IF SUPER^.Step(981,TRUE,'Step number 981') THEN		
	SUPER^.StepCompleteWhen((_runOneStep OR _runAllSteps) AND _finishStep);	
	IF _runOneStep THEN	
		_runOneStep := FALSE;
		RETURN;
	END_IF	
END_IF		
		
IF SUPER^.Step(982,TRUE,'Step number 982') THEN		
	SUPER^.StepCompleteWhen((_runOneStep OR _runAllSteps) AND _finishStep);	
	IF _runOneStep THEN	
		_runOneStep := FALSE;
		RETURN;
	END_IF	
END_IF		
		
IF SUPER^.Step(983,TRUE,'Step number 983') THEN		
	SUPER^.StepCompleteWhen((_runOneStep OR _runAllSteps) AND _finishStep);	
	IF _runOneStep THEN	
		_runOneStep := FALSE;
		RETURN;
	END_IF	
END_IF		
		
IF SUPER^.Step(984,TRUE,'Step number 984') THEN		
	SUPER^.StepCompleteWhen((_runOneStep OR _runAllSteps) AND _finishStep);	
	IF _runOneStep THEN	
		_runOneStep := FALSE;
		RETURN;
	END_IF	
END_IF		
		
IF SUPER^.Step(985,TRUE,'Step number 985') THEN		
	SUPER^.StepCompleteWhen((_runOneStep OR _runAllSteps) AND _finishStep);	
	IF _runOneStep THEN	
		_runOneStep := FALSE;
		RETURN;
	END_IF	
END_IF		
		
IF SUPER^.Step(986,TRUE,'Step number 986') THEN		
	SUPER^.StepCompleteWhen((_runOneStep OR _runAllSteps) AND _finishStep);	
	IF _runOneStep THEN	
		_runOneStep := FALSE;
		RETURN;
	END_IF	
END_IF		
		
IF SUPER^.Step(987,TRUE,'Step number 987') THEN		
	SUPER^.StepCompleteWhen((_runOneStep OR _runAllSteps) AND _finishStep);	
	IF _runOneStep THEN	
		_runOneStep := FALSE;
		RETURN;
	END_IF	
END_IF		
		
IF SUPER^.Step(988,TRUE,'Step number 988') THEN		
	SUPER^.StepCompleteWhen((_runOneStep OR _runAllSteps) AND _finishStep);	
	IF _runOneStep THEN	
		_runOneStep := FALSE;
		RETURN;
	END_IF	
END_IF		
		
IF SUPER^.Step(989,TRUE,'Step number 989') THEN		
	SUPER^.StepCompleteWhen((_runOneStep OR _runAllSteps) AND _finishStep);	
	IF _runOneStep THEN	
		_runOneStep := FALSE;
		RETURN;
	END_IF	
END_IF		
		
IF SUPER^.Step(990,TRUE,'Step number 990') THEN		
	SUPER^.StepCompleteWhen((_runOneStep OR _runAllSteps) AND _finishStep);	
	IF _runOneStep THEN	
		_runOneStep := FALSE;
		RETURN;
	END_IF	
END_IF		
		
IF SUPER^.Step(991,TRUE,'Step number 991') THEN		
	SUPER^.StepCompleteWhen((_runOneStep OR _runAllSteps) AND _finishStep);	
	IF _runOneStep THEN	
		_runOneStep := FALSE;
		RETURN;
	END_IF	
END_IF		
		
IF SUPER^.Step(992,TRUE,'Step number 992') THEN		
	SUPER^.StepCompleteWhen((_runOneStep OR _runAllSteps) AND _finishStep);	
	IF _runOneStep THEN	
		_runOneStep := FALSE;
		RETURN;
	END_IF	
END_IF		
		
IF SUPER^.Step(993,TRUE,'Step number 993') THEN		
	SUPER^.StepCompleteWhen((_runOneStep OR _runAllSteps) AND _finishStep);	
	IF _runOneStep THEN	
		_runOneStep := FALSE;
		RETURN;
	END_IF	
END_IF		
		
IF SUPER^.Step(994,TRUE,'Step number 994') THEN		
	SUPER^.StepCompleteWhen((_runOneStep OR _runAllSteps) AND _finishStep);	
	IF _runOneStep THEN	
		_runOneStep := FALSE;
		RETURN;
	END_IF	
END_IF		
		
IF SUPER^.Step(995,TRUE,'Step number 995') THEN		
	SUPER^.StepCompleteWhen((_runOneStep OR _runAllSteps) AND _finishStep);	
	IF _runOneStep THEN	
		_runOneStep := FALSE;
		RETURN;
	END_IF	
END_IF		
		
IF SUPER^.Step(996,TRUE,'Step number 996') THEN		
	SUPER^.StepCompleteWhen((_runOneStep OR _runAllSteps) AND _finishStep);	
	IF _runOneStep THEN	
		_runOneStep := FALSE;
		RETURN;
	END_IF	
END_IF		
		
IF SUPER^.Step(997,TRUE,'Step number 997') THEN		
	SUPER^.StepCompleteWhen((_runOneStep OR _runAllSteps) AND _finishStep);	
	IF _runOneStep THEN	
		_runOneStep := FALSE;
		RETURN;
	END_IF	
END_IF		
		
IF SUPER^.Step(998,TRUE,'Step number 998') THEN		
	SUPER^.StepCompleteWhen((_runOneStep OR _runAllSteps) AND _finishStep);	
	IF _runOneStep THEN	
		_runOneStep := FALSE;
		RETURN;
	END_IF	
END_IF		
		
IF SUPER^.Step(999,TRUE,'Step number 999') THEN		
	SUPER^.StepCompleteWhen((_runOneStep OR _runAllSteps) AND _finishStep);	
	IF _runOneStep THEN	
		_runOneStep := FALSE;
		RETURN;
	END_IF	
END_IF		
		
IF SUPER^.Step(1000,TRUE,'Step number 1000') THEN		
	SUPER^.StepCompleteWhen((_runOneStep OR _runAllSteps) AND _finishStep);	
	IF _runOneStep THEN	
		_runOneStep := FALSE;
		RETURN;
	END_IF	
END_IF		
		
IF SUPER^.Step(1001,TRUE,'Step number 1001') THEN		
	SUPER^.StepCompleteWhen((_runOneStep OR _runAllSteps) AND _finishStep);	
	IF _runOneStep THEN	
		_runOneStep := FALSE;
		RETURN;
	END_IF	
END_IF		
		
IF SUPER^.Step(1002,TRUE,'Step number 1002') THEN		
	SUPER^.StepCompleteWhen((_runOneStep OR _runAllSteps) AND _finishStep);	
	IF _runOneStep THEN	
		_runOneStep := FALSE;
		RETURN;
	END_IF	
END_IF		
		
IF SUPER^.Step(1003,TRUE,'Step number 1003') THEN		
	SUPER^.StepCompleteWhen((_runOneStep OR _runAllSteps) AND _finishStep);	
	IF _runOneStep THEN	
		_runOneStep := FALSE;
		RETURN;
	END_IF	
END_IF		
		
IF SUPER^.Step(1004,TRUE,'Step number 1004') THEN		
	SUPER^.StepCompleteWhen((_runOneStep OR _runAllSteps) AND _finishStep);	
	IF _runOneStep THEN	
		_runOneStep := FALSE;
		RETURN;
	END_IF	
END_IF		
		
IF SUPER^.Step(1005,TRUE,'Step number 1005') THEN		
	SUPER^.StepCompleteWhen((_runOneStep OR _runAllSteps) AND _finishStep);	
	IF _runOneStep THEN	
		_runOneStep := FALSE;
		RETURN;
	END_IF	
END_IF		
		
IF SUPER^.Step(1006,TRUE,'Step number 1006') THEN		
	SUPER^.StepCompleteWhen((_runOneStep OR _runAllSteps) AND _finishStep);	
	IF _runOneStep THEN	
		_runOneStep := FALSE;
		RETURN;
	END_IF	
END_IF		
		
IF SUPER^.Step(1007,TRUE,'Step number 1007') THEN		
	SUPER^.StepCompleteWhen((_runOneStep OR _runAllSteps) AND _finishStep);	
	IF _runOneStep THEN	
		_runOneStep := FALSE;
		RETURN;
	END_IF	
END_IF		
		
IF SUPER^.Step(1008,TRUE,'Step number 1008') THEN		
	SUPER^.StepCompleteWhen((_runOneStep OR _runAllSteps) AND _finishStep);	
	IF _runOneStep THEN	
		_runOneStep := FALSE;
		RETURN;
	END_IF	
END_IF		
		
IF SUPER^.Step(1009,TRUE,'Step number 1009') THEN		
	SUPER^.StepCompleteWhen((_runOneStep OR _runAllSteps) AND _finishStep);	
	IF _runOneStep THEN	
		_runOneStep := FALSE;
		RETURN;
	END_IF	
END_IF		
		
IF SUPER^.Step(1010,TRUE,'Step number 1010') THEN		
	SUPER^.StepCompleteWhen((_runOneStep OR _runAllSteps) AND _finishStep);	
	IF _runOneStep THEN	
		_runOneStep := FALSE;
		RETURN;
	END_IF	
END_IF		
		
IF SUPER^.Step(1011,TRUE,'Step number 1011') THEN		
	SUPER^.StepCompleteWhen((_runOneStep OR _runAllSteps) AND _finishStep);	
	IF _runOneStep THEN	
		_runOneStep := FALSE;
		RETURN;
	END_IF	
END_IF		
		
IF SUPER^.Step(1012,TRUE,'Step number 1012') THEN		
	SUPER^.StepCompleteWhen((_runOneStep OR _runAllSteps) AND _finishStep);	
	IF _runOneStep THEN	
		_runOneStep := FALSE;
		RETURN;
	END_IF	
END_IF		
		
IF SUPER^.Step(1013,TRUE,'Step number 1013') THEN		
	SUPER^.StepCompleteWhen((_runOneStep OR _runAllSteps) AND _finishStep);	
	IF _runOneStep THEN	
		_runOneStep := FALSE;
		RETURN;
	END_IF	
END_IF		
		
IF SUPER^.Step(1014,TRUE,'Step number 1014') THEN		
	SUPER^.StepCompleteWhen((_runOneStep OR _runAllSteps) AND _finishStep);	
	IF _runOneStep THEN	
		_runOneStep := FALSE;
		RETURN;
	END_IF	
END_IF		
		
IF SUPER^.Step(1015,TRUE,'Step number 1015') THEN		
	SUPER^.StepCompleteWhen((_runOneStep OR _runAllSteps) AND _finishStep);	
	IF _runOneStep THEN	
		_runOneStep := FALSE;
		RETURN;
	END_IF	
END_IF		
		
IF SUPER^.Step(1016,TRUE,'Step number 1016') THEN		
	SUPER^.StepCompleteWhen((_runOneStep OR _runAllSteps) AND _finishStep);	
	IF _runOneStep THEN	
		_runOneStep := FALSE;
		RETURN;
	END_IF	
END_IF		
		
IF SUPER^.Step(1017,TRUE,'Step number 1017') THEN		
	SUPER^.StepCompleteWhen((_runOneStep OR _runAllSteps) AND _finishStep);	
	IF _runOneStep THEN	
		_runOneStep := FALSE;
		RETURN;
	END_IF	
END_IF		
		
IF SUPER^.Step(1018,TRUE,'Step number 1018') THEN		
	SUPER^.StepCompleteWhen((_runOneStep OR _runAllSteps) AND _finishStep);	
	IF _runOneStep THEN	
		_runOneStep := FALSE;
		RETURN;
	END_IF	
END_IF		
		
IF SUPER^.Step(1019,TRUE,'Step number 1019') THEN		
	SUPER^.StepCompleteWhen((_runOneStep OR _runAllSteps) AND _finishStep);	
	IF _runOneStep THEN	
		_runOneStep := FALSE;
		RETURN;
	END_IF	
END_IF		
		
IF SUPER^.Step(1020,TRUE,'Step number 1020') THEN		
	SUPER^.StepCompleteWhen((_runOneStep OR _runAllSteps) AND _finishStep);	
	IF _runOneStep THEN	
		_runOneStep := FALSE;
		RETURN;
	END_IF	
END_IF		
		
IF SUPER^.Step(1021,TRUE,'Step number 1021') THEN		
	SUPER^.StepCompleteWhen((_runOneStep OR _runAllSteps) AND _finishStep);	
	IF _runOneStep THEN	
		_runOneStep := FALSE;
		RETURN;
	END_IF	
END_IF		
		
IF SUPER^.Step(1022,TRUE,'Step number 1022') THEN		
	SUPER^.StepCompleteWhen((_runOneStep OR _runAllSteps) AND _finishStep);	
	IF _runOneStep THEN	
		_runOneStep := FALSE;
		RETURN;
	END_IF	
END_IF		
		
IF SUPER^.Step(1023,TRUE,'Step number 1023') THEN		
	SUPER^.StepCompleteWhen((_runOneStep OR _runAllSteps) AND _finishStep);	
	IF _runOneStep THEN	
		_runOneStep := FALSE;
		RETURN;
	END_IF	
END_IF		
		
//******************************************************************
IF SUPER^.Step(_stepId,_enabled,_stepDescription) THEN
	SUPER^.StepCompleteWhen((_runOneStep OR _runAllSteps) AND _finishStep);	
	IF _runOneStep THEN	
		_runOneStep := FALSE;
		RETURN;
	END_IF		
END_IF
END_METHOD

METHOD PROTECTED OnSequenceCompleted
_onSequenceCompleteCount := _onSequenceCompleteCount + 1;
END_METHOD

METHOD PROTECTED OnSequencerError
VAR_INPUT
	inErrorId : eSequencerError;
END_VAR
CASE inErrorId OF
	eSequencerError.noError :
		_onSequencerErrorCount := _onSequencerErrorCount + 0;
	eSequencerError.NotUniqueStepId :
		_onSequencerErrorCount := _onSequencerErrorCount + 10;
	eSequencerError.StepIdHasBeenChanged :
		_onSequencerErrorCount := _onSequencerErrorCount + 20;
	eSequencerError.OrderOfTheStepHasBeenChanged :
		_onSequencerErrorCount := _onSequencerErrorCount + 40;
	eSequencerError.StepWithRequestedIdDoesNotExists :
		_onSequencerErrorCount := _onSequencerErrorCount + 50;
	eSequencerError.MultipleRequestStepMethodCall :
		_onSequencerErrorCount := _onSequencerErrorCount + 60;
	eSequencerError.StepIdTooLow :
		_onSequencerErrorCount := _onSequencerErrorCount + 70;
	eSequencerError.StepIdTooHigh :
		_onSequencerErrorCount := _onSequencerErrorCount + 80;
	ELSE
		_onSequencerErrorCount := _onSequencerErrorCount + 0;
END_CASE
END_METHOD

METHOD PROTECTED OnStateChange
VAR_INPUT
	PreviousState	: INT;
	NewState 		: INT;
END_VAR
THIS^._onStateChangeCount := THIS^._onStateChangeCount + 1;

_stateChangeFrom := PreviousState;
_stateChangeTo := NewState;

IF _callRestoreInOnStateChange THEN
	Restore();
END_IF
END_METHOD

METHOD PROTECTED OnStepCompleted
_onCompleteStepCount := _onCompleteStepCount + 1;
END_METHOD

PROPERTY INTERNAL RequestStepCycle : UINT
GET
RequestStepCycle := _requestStepCycle;
END_GET
SET
_requestStepCycle := RequestStepCycle;
END_SET
END_PROPERTY

METHOD INTERNAL SequencerClose
SUPER^._Close();
END_METHOD

METHOD INTERNAL SequencerHasError : BOOL
SequencerHasError := SUPER^._sequencerHasError;
END_METHOD

METHOD INTERNAL SequencerOpen
SUPER^._Open();
END_METHOD

METHOD INTERNAL SetChildState 
VAR_INPUT
	inState			:	INT;
END_VAR
THIS^._myTcoState.ChangeState(inState);
END_METHOD

METHOD INTERNAL SetCurrentStep 
VAR_INPUT
	inStepID 			:	INT;
	inStepDescription	:	STRING(254);
END_VAR
THIS^._currentStep.ID			:=	inStepID;
THIS^._currentStep.Description	:=	inStepDescription;
END_METHOD

METHOD SetCurrentStepToErrorState : BOOL
_currentStep.Status := TcoCore.eStepStatus.Error;

SetCurrentStepToErrorState := _currentStep.Status = TcoCore.eStepStatus.Error;
END_METHOD

METHOD SetCyclicMode : BOOL
ModeController.Mode := eSequencerMode.CyclicMode;

SetCyclicMode := ModeController.Mode = eSequencerMode.CyclicMode;
END_METHOD

METHOD SetInvalidMode : BOOL
ModeController.Mode := eSequencerMode.Invalid;

SetInvalidMode := ModeController.Mode = eSequencerMode.Invalid;
END_METHOD

METHOD INTERNAL SetNumberOfSteps 
VAR_INPUT
	inNumberOfSteps : UINT;
END_VAR
_stepCounter 						:=	inNumberOfSteps;
_numberOfStepsInSequence			:=	inNumberOfSteps;
_previousNumberOfStepsInSequence 	:=	inNumberOfSteps;
END_METHOD

METHOD INTERNAL SetSequenceAsChecked
_stepIDUniquenessChecked := TRUE;
_StepIdUniquenessControlState := eStepIdUniquenessControlState.Done;
END_METHOD

METHOD INTERNAL SetSequenceAsNotChecked
_stepIDUniquenessChecked := FALSE;
_StepIdUniquenessControlState := eStepIdUniquenessControlState.NotYetStarted;
END_METHOD

METHOD SetStepMode : BOOL
ModeController.Mode := eSequencerMode.StepMode;

SetStepMode := ModeController.Mode = eSequencerMode.StepMode;
END_METHOD

METHOD INTERNAL SetTestParams
VAR_INPUT
	inRunOneStep		:	BOOL;
	inRunAllSteps		:	BOOL;
	inFinishStep		:	BOOL;
	inID				:	UINT;
	inEnabled			:	BOOL;
	inStepDescription	:	STRING(254);	
END_VAR
THIS^._runOneStep		:=			inRunOneStep;
THIS^._runAllSteps 		:= 			inRunAllSteps;
THIS^._finishStep 		:= 			inFinishStep;
THIS^._stepId 				:=			inID;
THIS^._enabled 			:= 			inEnabled;
THIS^._stepDescription 	:=			inStepDescription;
END_METHOD

METHOD StepCount 
VAR_INPUT
    inTotalStepNumber : UINT;
    inFinishStep : BOOL;
END_VAR
VAR 
	i : INT;
	_lastStepId : INT;
END_VAR
FOR i:=0 TO inTotalStepNumber DO
	IF SUPER^.Step(i,TRUE,CONCAT('Step number ',INT_TO_STRING(i))) THEN		
		SUPER^.StepCompleteWhen(inFinishStep);	
	END_IF	
END_FOR
END_METHOD

{attribute 'TcRpcEnable'}
METHOD INTERNAL UpdateCurrentStepDetails
_currentStepId				:=	SUPER^._currentStep.ID;
_currentStepOrder			:=	SUPER^._currentStep.Order;
_currentStepEnabled			:=	SUPER^._currentStep.Enabled;
_currentStepDescription		:=	SUPER^._currentStep.Description;
_currentStepStatus			:=	SUPER^._currentStep.Status;
_currentStepDuration		:=	SUPER^._currentStep.Duration;
END_METHOD

END_FUNCTION_BLOCK

(* stored: Version 1.1.0.1
   POU _TcoSequencer: Id {ac19fe4f-0c0e-08e9-3df5-0840192e4ee2}, SpecialFunc None
   Folder _Tests: Id {36ff3928-274d-02d5-18e6-23dcd25a0584}
   Method _RequestStep: Id {7aa88188-6d52-03a0-2257-f5ace3c373f6}
   Method _SequenceComplete: Id {bb57ddc4-708a-0b87-2b40-163e4ea27d45}
   Method _Step: Id {9a6df11c-2565-03db-3c82-b0919c6a6202}
   Method _StepBackward: Id {bb6fa187-eb1c-0571-2358-79713c7a9719}
   Method _StepCompleteWhen: Id {e0d9eb39-b1b6-0ab0-0c06-820f1dca6b2f}
   Method _StepForward: Id {27ff14c0-bd91-0858-2810-1f7c5fd2dc67}
   Method _StepIn: Id {00d65f73-93ab-04a1-31ca-6a19a3e4c8dd}
   Method ChildHasAutoRestoreEnabled: Id {2fe344f3-4fea-0846-0ec8-378fe51cb4c6}
   Method ChildIsAutoRestorable: Id {e0cb2365-b187-0b05-2101-33f128967786}
   Method CleanupPointers: Id {c754833e-788e-0dc0-39b2-57f91228c555}
   Method ClearNumberOfSteps: Id {ccb8339d-f888-01c2-334c-f78620010950}
   Method GetChildState: Id {aaac1bd4-eac0-002e-3f58-ea6c5e49e949}
   Method GetNumberOfStepsInSequence: Id {154b9cc4-fcc7-08ab-0ee3-cde964c24006}
   Method GetSequencerErrorId: Id {cfa5c7b8-bdaa-0dc9-318b-07d87a737808}
   Method GetTextOfTheMostImportantMessage: Id {0f5e0607-86a0-04f2-3053-f70b778527fb}
   Method HasAutoRestoreEnabled: Id {13163512-5f77-0a1f-15bd-0485ab98dc6e}
   Method IsAutoRestorable: Id {78b773c3-e01b-01ec-3871-0a0bdbd810d6}
   Method IsFirstStepEntry: Id {4f006540-c701-07be-1eb3-95b9c8a360ee}
   Method Main: Id {3a6cbc53-5690-0480-174f-e4140d338a45}
   Method OnSequenceCompleted: Id {2fd78922-07d4-01ec-1736-1c3b4b7d9bd8}
   Method OnSequencerError: Id {812d3e89-fa98-0c05-2d57-bd1b9d1501be}
   Method OnStateChange: Id {a3a0e1a2-27bc-0384-1d2b-01018017d7b0}
   Method OnStepCompleted: Id {154d4f23-050b-01f6-08b9-2a631c3ec621}
   Property RequestStepCycle: Id {c2da0157-c6b1-052f-064f-3e3f6d17de69}
   Get Get: Id {6b43bca9-2a6f-0436-073d-241b14a17d9a}
   Set Set: Id {66bd96b6-e8a3-0fe0-344b-3b831339bba2}
   Method SequencerClose: Id {f3addcb4-0fda-0a2d-0925-430c6f4ad3f8}
   Method SequencerHasError: Id {07e19515-04c8-048f-12a4-f42415093577}
   Method SequencerOpen: Id {b4334737-6cb3-0eba-0d2f-cd067be7b53d}
   Method SetChildState: Id {60024768-516f-0fd2-2f16-e270836f2db6}
   Method SetCurrentStep: Id {223d2a4f-ee82-0c54-0227-548f61243f4d}
   Method SetCurrentStepToErrorState: Id {5c3befd4-bb7c-0fc8-2440-5e08fffd4f9e}
   Method SetCyclicMode: Id {d046251b-754e-073d-2a86-854f5889d9d0}
   Method SetInvalidMode: Id {9fac0342-f3de-0c15-053d-bbfecf3074ce}
   Method SetNumberOfSteps: Id {a8a0d4fb-e225-0fb8-3c9b-d2a796c1b2ec}
   Method SetSequenceAsChecked: Id {43e68eca-b921-0c50-2ca5-03882ac05b27}
   Method SetSequenceAsNotChecked: Id {09a6a7e6-7763-040e-016a-fc5c2ce30618}
   Method SetStepMode: Id {03d14d20-a375-0456-1afe-147a68ccc6ff}
   Method SetTestParams: Id {7a624c26-ee8b-0b24-15f9-09fad6ccc521}
   Method StepCount: Id {04d7f514-94fe-03d1-1b6f-5300a828c9d4}
   Method UpdateCurrentStepDetails: Id {590d6a94-7182-0c50-1bd0-bf34e87df18c} *)
